(*
SPDX-FileCopyrightText: c 2026 Oleksandr Tiutyk <trofimich@gmail.com>
SPDX-License-Identifier: MIT
License: https://opensource.org/license/mit
*)

(*!
<summary>Checks stable membership for raw and generic matching and missing values.</summary>
<description>
Borrows one group-owned set reserved for this case. Use from one task at a stable address.
Teardown clears the set and releases its owned entries before publication.
</description>
*)

{attribute 'no_assign'}
{attribute 'no_explicit_call' := 'do not call this function block directly'}
FUNCTION_BLOCK UniqueDataSetContainsTest EXTENDS TOF_Testing.SingleCycleTest
VAR_STAT
	{attribute 'hide'}
	_ClassName : STRING := __POUNAME();
END_VAR
VAR
	_Set : TOF_Collections.IUniqueDataSet;
END_VAR

(*!
<summary>Clears the fixture before the runner publishes the result.</summary>
<description>
Also runs after an unexpected exception interrupts the case.
</description>
*)
METHOD PROTECTED AfterTest
_Set.Clear();
END_METHOD

//! <summary>Borrows the concrete class name. Callers must not modify it.</summary>
{attribute 'monitoring' := 'call'}
PROPERTY ClassName : REFERENCE TO STRING
GET
ClassName REF= _ClassName;
END_GET
END_PROPERTY

(*!
<summary>Checks stable membership for raw and generic matching and missing values.</summary>
*)
METHOD PROTECTED ExecuteTest
VAR
	values : ARRAY [0..6] OF STRING :=
		['String0', 'String1', 'String2', 'String3', 'String4', 'String5', 'String6'];
	i : DINT;
	missingValue : STRING := 'String9';
	query : TOF_Core.GENERIC_VALUE;
END_VAR
FOR i := 6 TO 0 BY -1 DO
	_Set.SetCopy(value := values[i]);
END_FOR

Assert.ThatBool(
	actual := _Set.Contains(value := values[3]),
	message := "Contains must find a stored value"
).IsTrue();

Assert.ThatBool(
	actual := _Set.Contains(value := missingValue),
	message := "Contains must reject an absent value"
).IsFalse();

query := TOF_Core.GenericValueFactory.FromStringReference(value := values[3]);
Assert.ThatBool(
	actual := _Set.ContainsGeneric(value := query, releaseValue := FALSE),
	message := "ContainsGeneric must find a stored value"
).IsTrue();

query := TOF_Core.GenericValueFactory.FromStringReference(value := missingValue);
Assert.ThatBool(
	actual := _Set.ContainsGeneric(value := query, releaseValue := FALSE),
	message := "ContainsGeneric must reject an absent value"
).IsFalse();

Assert.ThatDInt(
	actual := _Set.Length,
	message := "Lookup must preserve all seven entries"
).ToBe(expected := DINT#7);
END_METHOD

(*!
<summary>Binds the unique set fixture for this case.</summary>
<description>
Stores a borrowed interface without invoking the fixture. The owning group keeps it alive and
reserves it for this case. TestElement initializes the name and parent.
</description>
<param name="name">Display name of this case.</param>
<param name="parent">Group that owns this case.</param>
<param name="dataSet">Required live unique set reserved for this case.</param>
*)
METHOD FB_init : BOOL
VAR_INPUT
	bInitRetains: BOOL; // TRUE: the retain variables are initialized (reset warm / reset cold)
	bInCopyCode: BOOL; // TRUE: the instance will be copied to the copy code afterward (online change)
	name : WSTRING;
	parent : TOF_Testing.ITestElement;
	dataSet : TOF_Collections.IUniqueDataSet;
END_VAR
_Set := dataSet;
FB_init := TRUE;
END_METHOD

//! <summary>Borrows the compiler-initialized namespace name. Callers must not modify it.</summary>
{attribute 'monitoring' := 'call'}
PROPERTY NamespaceName : REFERENCE TO STRING
GET
NamespaceName REF= CurrentNamespace.Name;
END_GET
END_PROPERTY

//! <summary>Reports the concrete instance size in bytes.</summary>
{attribute 'monitoring' := 'call'}
PROPERTY SelfSize : ULINT
GET
SelfSize := XSIZEOF(THIS^);
END_GET
END_PROPERTY

END_FUNCTION_BLOCK

(* stored: Version 1.1.0.1, ProductVersion 3.1.4026.21
   POU UniqueDataSetContainsTest: Id {59f51ea0-e39e-4d6e-a4c3-0feebb775300}, SpecialFunc None
   Method AfterTest: Id {344a2be2-d5e4-4524-9db4-5d6eda55859e}
   Property ClassName: Id {7f5cc86b-b79e-4235-9d08-75fb588a113b}
   Get Get: Id {05d5c265-deeb-4f27-b063-ae39e1534258}
   Method ExecuteTest: Id {c48bfafb-ba19-4b24-b910-5a36794ce3b0}
   Method FB_init: Id {9d2a28a5-ee67-4b43-8a1b-4edebcf5cfd9}
   Property NamespaceName: Id {d9338d1c-d3c3-452c-bcd4-aa8097a7d542}
   Get Get: Id {b769c79e-010e-4868-8639-4ee0d3d823f5}
   Property SelfSize: Id {12fda590-7b2d-4906-913c-5dee5079ef23}
   Get Get: Id {2f25ccf6-fd69-44b0-8905-a0a87539815e} *)
